Fanuc KAREL source: KA00104.KL

PROGRAM KA00104
%NOLOCKGROUP
VAR
  SRC: VECTOR
  DST: JOINTPOS
BEGIN
  SRC.X = 1.0
  DST = SRC
END KA00104
